// TwinCAT 3 PLC project TwinCAT_OpenFramework_HowTo
// Title: TwinCAT Open Framework HowTo
// Company: Oleksandr Tiutyk FOP
// Author: Oleksandr Tiutyk
// ProjectVersion: 1.0.13.0
// Description: Small samples how to use TwinCAT.OpenFramework
// ProgramVersion: 3.1.4026.28
// libraries:
//   [TwinCAT Open Framework Testing], * (Oleksandr Tiutyk FOP)
//   [TwinCAT Open Framework Core], * (Oleksandr Tiutyk FOP)
//   [TwinCAT Open Framework IO Models], * (Oleksandr Tiutyk FOP)
//   Tc2_Standard, * (Beckhoff Automation GmbH)
//   Tc2_System, * (Beckhoff Automation GmbH)
// project tree:
//   / CurrentNamespace.TcGVL, MAIN.TcPOU, PlcTask.TcTTO
//   Testing/ AdditionTestRunner.TcPOU, BasicTestRunner.TcPOU, TimerDelayTestRunner.TcPOU, AdditionTest.TcPOU, TimerDelayTest.TcPOU, SingleCycleTestExample.TcPOU, MultiCycleTestExample.TcPOU, TimingTestGroup.TcPOU, BasicTestGroup.TcPOU, GroupedTestExample.TcPOU
//   IO/ IOModelsExample.TcPOU
//   Version/ Global_Version.TcGVL
// (motion and I/O tree: see PLC project twincat_openframework_core)
// real-time tasks:
//   TASK PlcTask: cycle T#10ms, priority 20, ADS port 350
//   TASK TestTask: cycle T#10ms, priority 1, ADS port 351
//   TASK RunnerTestTask: cycle T#10ms, priority 2, ADS port 354
//   TASK HowToTask: cycle T#10ms, priority 22, ADS port 353
// variable links:

CONFIGURATION TwinCAT_OpenFramework_HowTo
    RESOURCE PLC ON TwinCAT3
        TASK PlcTask(INTERVAL := T#10ms, PRIORITY := 22);
        PROGRAM MAIN WITH PlcTask : MAIN;
    END_RESOURCE
END_CONFIGURATION

// ---- CurrentNamespace.TcGVL
(*
SPDX-FileCopyrightText: © 2026 Oleksandr Tiutyk <trofimich@gmail.com>
SPDX-License-Identifier: MIT
License: https://opensource.org/license/mit
*)

{attribute 'qualified_only'}
VAR_GLOBAL
	Name : STRING := 'TOF_Tests';
END_VAR

// ---- Version/Global_Version.TcGVL
{attribute 'TcGenerated'}
{attribute 'no-analysis'}
{attribute 'linkalways'}
// This function has been automatically generated from the project information.
VAR_GLOBAL CONSTANT
	{attribute 'const_non_replaced'}
	stLibVersion_TwinCAT_Open_Framework_HowTo : ST_LibVersion := (iMajor := 1, iMinor := 0, iBuild := 13, iRevision := 0, nFlags := 0, sVersion := '1.0.13.0');
END_VAR

// ---- MAIN.TcPOU
(*
SPDX-FileCopyrightText: © 2026 Oleksandr Tiutyk <trofimich@gmail.com>
SPDX-License-Identifier: MIT
License: https://opensource.org/license/mit
*)

(*!
<summary>Runs the standalone single-cycle testing example through its explicit execution method.</summary>
<description>Mapped by PlcTask. Do not also map SingleCycleTestExample to a task while this entry is used.</description>
*)

{attribute 'no_explicit_call' := 'do not call this function block directly'}
PROGRAM MAIN
VAR
	{attribute 'hide'}
	_ClassName : STRING := __POUNAME();
END_VAR

SingleCycleTestExample.Execute();

(*!
<summary>Borrows the concrete program name for its lifetime.</summary>
<description>Borrowed read-only storage; callers must not modify it.</description>
*)
{attribute 'monitoring' := 'call'}
PROPERTY ClassName : REFERENCE TO STRING
GET
ClassName REF= _ClassName;
END_GET
END_PROPERTY

(*!
<summary>Borrows the project namespace for the program lifetime.</summary>
<description>Borrowed read-only storage; callers must not modify it.</description>
*)
{attribute 'monitoring' := 'call'}
PROPERTY NamespaceName : REFERENCE TO STRING
GET
NamespaceName REF= CurrentNamespace.Name;
END_GET
END_PROPERTY

END_PROGRAM

// ---- Testing/SingleCycleTestExample.TcPOU
(*
SPDX-FileCopyrightText: © 2026 Oleksandr Tiutyk <trofimich@gmail.com>
SPDX-License-Identifier: MIT
License: https://opensource.org/license/mit
*)

(*!
<summary>Runs one single-cycle test directly, without a group.</summary>
<description>
Map this program to one cyclic PLC task or call its Execute method once per cycle from that task.
The concrete runner owns the tests; the program owns the reporter and performs task
cleanup at the end of every scan. Inspect _Runner.IsFinished, AllPassed and counts, then _Report.IsReady.
For independent task execution, assign SingleCycleTestExample and MultiCycleTestExample to different tasks.
They share no instances or mutable buffers. Do not assign the same program instance to multiple tasks.
</description>
*)

{attribute 'no_explicit_call' := 'do not call this function block directly'}
PROGRAM SingleCycleTestExample
VAR
	{attribute 'hide'}
	_ClassName : STRING := __POUNAME();

	_Runner : AdditionTestRunner;
	_Report : TOF_Testing.JUnitXmlReporter;
	_Configured : BOOL;
END_VAR

Execute();

//! <summary>Borrows the concrete program name for its lifetime; callers must not modify it.</summary>
{attribute 'monitoring' := 'call'}
PROPERTY ClassName : REFERENCE TO STRING
GET
ClassName REF= _ClassName;
END_GET
END_PROPERTY

(*!
<summary>Advances this example and performs standalone task-boundary memory cleanup.</summary>
<description>
Call once per cycle from the owning task, either through this method or by mapping this PROGRAM to that task.
Do not drive both entry paths or share the instance between tasks. Use as the standalone example in its task;
hosts with additional transient-exception consumers must provide a shared boundary instead.
</description>
*)
METHOD Execute
IF NOT _Configured THEN
	_Runner.Reporter := _Report;
	_Configured := TRUE;
END_IF

_Runner.Execute(cleanupTaskMemory := TRUE);
END_METHOD

(*!
<summary>Provides the library namespace used in diagnostics.</summary>
<description>
Borrowed read-only reference to the compiler-initialized library namespace; no ownership transfer.
</description>
*)
{attribute 'monitoring' := 'call'}
PROPERTY NamespaceName : REFERENCE TO STRING
GET
NamespaceName REF= CurrentNamespace.Name;
END_GET
END_PROPERTY

END_PROGRAM

// ---- Testing/AdditionTestRunner.TcPOU
(*
SPDX-License-Identifier: MIT
License: https://opensource.org/license/mit
*)

(*!
<summary>Runs one owned addition test without a group.</summary>
<description>
Owns persistent root instances and fixed child storage. Use from one task without reentry.
Children borrows the same array for the instance lifetime. Root parents remain zero.
</description>
*)

{attribute 'no_assign'}
{attribute 'no_explicit_call' := 'do not call this function block directly'}
FUNCTION_BLOCK AdditionTestRunner EXTENDS TOF_Testing.TestRunner<1>
VAR_STAT
	//! <summary>Class name shared by instances of this concrete runner.</summary>
	{attribute 'hide'}
	_ClassName : STRING := __POUNAME();
END_VAR
VAR
	{attribute 'hide'}
	{attribute 'init_namespace'}
	_NamespaceName : STRING;
END_VAR
VAR_OUTPUT
	//! <summary>Owned root element used by this runner.</summary>
	Root : AdditionTest(name := "Addition", parent := 0);
END_VAR
VAR
	_Children : ARRAY [0.._ChildCount - 1] OF TOF_Testing.ITestElement :=
	[
		Root
	];
END_VAR

(*!
<summary>Borrows the concrete class name; callers must not modify the returned storage.</summary>
*)
{attribute 'monitoring' := 'call'}
PROPERTY ClassName : REFERENCE TO STRING
GET
ClassName REF= _ClassName;
END_GET
END_PROPERTY

(*!
<summary>Borrows the concrete namespace name for the instance lifetime; callers must not modify it.</summary>
*)
{attribute 'monitoring' := 'call'}
PROPERTY NamespaceName : REFERENCE TO STRING
GET
NamespaceName REF= _NamespaceName;
END_GET
END_PROPERTY

(*!
<summary>Reports the complete concrete instance size.</summary>
*)
{attribute 'monitoring' := 'call'}
PROPERTY SelfSize : ULINT
GET
SelfSize := XSIZEOF(THIS^);
END_GET
END_PROPERTY

(*!
<summary>Borrows the unchanged persistent root array; application code must not modify it.</summary>
*)
{attribute 'monitoring' := 'call'}
PROPERTY Children : REFERENCE TO ARRAY [0.._ChildCount - 1] OF TOF_Testing.ITestElement
GET
Children REF= _Children;
END_GET
END_PROPERTY

END_FUNCTION_BLOCK

// ---- Testing/AdditionTest.TcPOU
(*
SPDX-FileCopyrightText: © 2026 Oleksandr Tiutyk <trofimich@gmail.com>
SPDX-License-Identifier: MIT
License: https://opensource.org/license/mit
*)

(*!
<summary>Shows a complete single-cycle test body without guards or contexts.</summary>
*)

{attribute 'no_explicit_call' := 'do not call this function block directly'}
FUNCTION_BLOCK AdditionTest EXTENDS TOF_Testing.SingleCycleTest
VAR_STAT
	{attribute 'hide'}
	_ClassName : STRING := __POUNAME();
END_VAR

//! <summary>Borrows the concrete class name for the lifetime of this instance; callers must not modify it.</summary>
{attribute 'monitoring' := 'call'}
PROPERTY ClassName : REFERENCE TO STRING
GET
ClassName REF= _ClassName;
END_GET
END_PROPERTY

(*!
<summary>Checks an arithmetic result and completes automatically on return.</summary>
*)
METHOD PROTECTED ExecuteTest
Assert.ThatDInt(actual := 2 + 3).ToBe(expected := 5);
END_METHOD

//! <summary>Borrows the compiler-initialized namespace; callers must not modify the returned reference.</summary>
{attribute 'monitoring' := 'call'}
PROPERTY NamespaceName : REFERENCE TO STRING
GET
NamespaceName REF= CurrentNamespace.Name;
END_GET
END_PROPERTY

//! <summary>Reports the complete concrete instance size, excluding separately allocated storage.</summary>
{attribute 'monitoring' := 'call'}
PROPERTY SelfSize : ULINT
GET
SelfSize := XSIZEOF(THIS^);
END_GET
END_PROPERTY

END_FUNCTION_BLOCK

// ---- Testing/BasicTestRunner.TcPOU
(*
SPDX-License-Identifier: MIT
License: https://opensource.org/license/mit
*)

(*!
<summary>Runs the owned basic test group and its nested timing group.</summary>
<description>
Owns persistent root instances and fixed child storage. Use from one task without reentry.
Children borrows the same array for the instance lifetime. Root parents remain zero.
</description>
*)

{attribute 'no_assign'}
{attribute 'no_explicit_call' := 'do not call this function block directly'}
FUNCTION_BLOCK BasicTestRunner EXTENDS TOF_Testing.TestRunner<1>
VAR_STAT
	//! <summary>Class name shared by instances of this concrete runner.</summary>
	{attribute 'hide'}
	_ClassName : STRING := __POUNAME();
END_VAR
VAR
	{attribute 'hide'}
	{attribute 'init_namespace'}
	_NamespaceName : STRING;
END_VAR
VAR_OUTPUT
	//! <summary>Owned root element used by this runner.</summary>
	Root : BasicTestGroup(name := "Basic", parent := 0);
END_VAR
VAR
	_Children : ARRAY [0.._ChildCount - 1] OF TOF_Testing.ITestElement :=
	[
		Root
	];
END_VAR

(*!
<summary>Borrows the concrete class name; callers must not modify the returned storage.</summary>
*)
{attribute 'monitoring' := 'call'}
PROPERTY ClassName : REFERENCE TO STRING
GET
ClassName REF= _ClassName;
END_GET
END_PROPERTY

(*!
<summary>Borrows the concrete namespace name for the instance lifetime; callers must not modify it.</summary>
*)
{attribute 'monitoring' := 'call'}
PROPERTY NamespaceName : REFERENCE TO STRING
GET
NamespaceName REF= _NamespaceName;
END_GET
END_PROPERTY

(*!
<summary>Reports the complete concrete instance size.</summary>
*)
{attribute 'monitoring' := 'call'}
PROPERTY SelfSize : ULINT
GET
SelfSize := XSIZEOF(THIS^);
END_GET
END_PROPERTY

(*!
<summary>Borrows the unchanged persistent root array; application code must not modify it.</summary>
*)
{attribute 'monitoring' := 'call'}
PROPERTY Children : REFERENCE TO ARRAY [0.._ChildCount - 1] OF TOF_Testing.ITestElement
GET
Children REF= _Children;
END_GET
END_PROPERTY

END_FUNCTION_BLOCK

// ---- Testing/BasicTestGroup.TcPOU
(*
SPDX-License-Identifier: MIT
License: https://opensource.org/license/mit
*)

(*!
<summary>Owns an arithmetic test and a nested timing group.</summary>
<description>
Owns persistent child storage and fixed parent associations. Use in one task without reentry.
Children is borrowed and must not be modified by application code. Constructor callbacks are not used.
</description>
*)

{attribute 'no_assign'}
{attribute 'no_explicit_call' := 'do not call this function block directly'}
FUNCTION_BLOCK BasicTestGroup EXTENDS TOF_Testing.TestGroup<2>
VAR_STAT
	{attribute 'hide'}
	_ClassName : STRING := __POUNAME();
END_VAR
VAR
	_Addition : AdditionTest(name := "Addition", parent := THIS^);
	_Timing : TimingTestGroup(name := "Timing", parent := THIS^);

	_Children : ARRAY [0.._ChildCount - 1] OF TOF_Testing.ITestElement :=
	[
		_Addition,
		_Timing
	];
END_VAR

//! <summary>Borrows the fixed array of this concrete group; do not modify it.</summary>
{attribute 'monitoring' := 'call'}
PROPERTY Children : REFERENCE TO ARRAY [0.._ChildCount - 1] OF TOF_Testing.ITestElement
GET
Children REF= _Children;
END_GET
END_PROPERTY

//! <summary>Borrows the concrete class name for the lifetime of this instance; callers must not modify it.</summary>
{attribute 'monitoring' := 'call'}
PROPERTY ClassName : REFERENCE TO STRING
GET
ClassName REF= _ClassName;
END_GET
END_PROPERTY

//! <summary>Borrows the compiler-initialized namespace; callers must not modify the returned reference.</summary>
{attribute 'monitoring' := 'call'}
PROPERTY NamespaceName : REFERENCE TO STRING
GET
NamespaceName REF= CurrentNamespace.Name;
END_GET
END_PROPERTY

//! <summary>Reports the complete concrete instance size, excluding separately allocated storage.</summary>
{attribute 'monitoring' := 'call'}
PROPERTY SelfSize : ULINT
GET
SelfSize := XSIZEOF(THIS^);
END_GET
END_PROPERTY

END_FUNCTION_BLOCK

// ---- Testing/TimingTestGroup.TcPOU
(*
SPDX-License-Identifier: MIT
License: https://opensource.org/license/mit
*)

(*!
<summary>Owns a timer-delay test as a static group.</summary>
<description>
Owns persistent child storage and fixed parent associations. Use in one task without reentry.
Children is borrowed and must not be modified by application code. Constructor callbacks are not used.
</description>
*)

{attribute 'no_assign'}
{attribute 'no_explicit_call' := 'do not call this function block directly'}
FUNCTION_BLOCK TimingTestGroup EXTENDS TOF_Testing.TestGroup<1>
VAR_STAT
	//! <summary>Class name shared by all instances of this function block.</summary>
	{attribute 'hide'}
	_ClassName : STRING := __POUNAME();
END_VAR
VAR
	_Timer : TimerDelayTest(name := "Timer delay", parent := THIS^);

	_Children : ARRAY [0.._ChildCount - 1] OF TOF_Testing.ITestElement :=
	[
		_Timer
	];
END_VAR

//! <summary>Borrows the fixed array of this concrete group; do not modify it.</summary>
{attribute 'monitoring' := 'call'}
PROPERTY Children : REFERENCE TO ARRAY [0.._ChildCount - 1] OF TOF_Testing.ITestElement
GET
Children REF= _Children;
END_GET
END_PROPERTY

//! <summary>Borrows the concrete class name for the lifetime of this instance; callers must not modify it.</summary>
{attribute 'monitoring' := 'call'}
PROPERTY ClassName : REFERENCE TO STRING
GET
ClassName REF= _ClassName;
END_GET
END_PROPERTY

//! <summary>Borrows the compiler-initialized namespace; callers must not modify the returned reference.</summary>
{attribute 'monitoring' := 'call'}
PROPERTY NamespaceName : REFERENCE TO STRING
GET
NamespaceName REF= CurrentNamespace.Name;
END_GET
END_PROPERTY

//! <summary>Reports the complete concrete instance size, excluding separately allocated storage.</summary>
{attribute 'monitoring' := 'call'}
PROPERTY SelfSize : ULINT
GET
SelfSize := XSIZEOF(THIS^);
END_GET
END_PROPERTY

END_FUNCTION_BLOCK

// ---- Testing/TimerDelayTest.TcPOU
(*
SPDX-FileCopyrightText: © 2026 Oleksandr Tiutyk <trofimich@gmail.com>
SPDX-License-Identifier: MIT
License: https://opensource.org/license/mit
*)

(*!
<summary>Shows persistent state and explicit completion in a multi-cycle test.</summary>
<description>
The inherited one-second deadline bounds waiting for a twenty-millisecond timer.
</description>
*)

{attribute 'no_explicit_call' := 'do not call this function block directly'}
FUNCTION_BLOCK TimerDelayTest EXTENDS TOF_Testing.MultiCycleTest
VAR
	_Timer : Tc2_Standard.TON;
END_VAR
VAR_STAT
	//! <summary>Class name shared by all instances of this function block.</summary>
	{attribute 'hide'}
	_ClassName : STRING := __POUNAME();
END_VAR
VAR
	{attribute 'hide'}
	{attribute 'init_namespace'}
	_NamespaceName : STRING;
END_VAR

(*!
<summary>Resets the timer after completion or failure.</summary>
*)
METHOD PROTECTED AfterTest
_Timer(IN := FALSE, PT := T#20MS);
END_METHOD

(*!
<summary>Resets the timer before each run.</summary>
*)
METHOD PROTECTED BeforeTest
_Timer(IN := FALSE, PT := T#20MS);
END_METHOD

//! <summary>Borrows the concrete class name for the lifetime of this instance; callers must not modify it.</summary>
{attribute 'monitoring' := 'call'}
PROPERTY ClassName : REFERENCE TO STRING
GET
ClassName REF= _ClassName;
END_GET
END_PROPERTY

(*!
<summary>Advances the timer once and returns DONE after its delay.</summary>
*)
METHOD PROTECTED ExecuteTest : TOF_Testing.TEST_CYCLE_RESULT
_Timer(IN := TRUE, PT := T#20MS);

IF _Timer.Q THEN
	Assert.ThatTime(actual := _Timer.ET).IsGreaterThanOrEquals(expected := T#20MS);
	ExecuteTest := TOF_Testing.TEST_CYCLE_RESULT.DONE;
ELSE
	ExecuteTest := TOF_Testing.TEST_CYCLE_RESULT.BUSY;
END_IF
END_METHOD

//! <summary>Borrows the compiler-initialized namespace; callers must not modify the returned reference.</summary>
{attribute 'monitoring' := 'call'}
PROPERTY NamespaceName : REFERENCE TO STRING
GET
NamespaceName REF= CurrentNamespace.Name;
END_GET
END_PROPERTY

//! <summary>Reports the complete concrete instance size, excluding separately allocated storage.</summary>
{attribute 'monitoring' := 'call'}
PROPERTY SelfSize : ULINT
GET
SelfSize := XSIZEOF(THIS^);
END_GET
END_PROPERTY

END_FUNCTION_BLOCK

// ---- Testing/TimerDelayTestRunner.TcPOU
(*
SPDX-License-Identifier: MIT
License: https://opensource.org/license/mit
*)

(*!
<summary>Runs one owned multi-cycle timer test.</summary>
<description>
Owns persistent root instances and fixed child storage. Use from one task without reentry.
Children borrows the same array for the instance lifetime. Root parents remain zero.
</description>
*)

{attribute 'no_assign'}
{attribute 'no_explicit_call' := 'do not call this function block directly'}
FUNCTION_BLOCK TimerDelayTestRunner EXTENDS TOF_Testing.TestRunner<1>
VAR_STAT
	//! <summary>Class name shared by instances of this concrete runner.</summary>
	{attribute 'hide'}
	_ClassName : STRING := __POUNAME();
END_VAR
VAR
	{attribute 'hide'}
	{attribute 'init_namespace'}
	_NamespaceName : STRING;
END_VAR
VAR_OUTPUT
	//! <summary>Owned root element used by this runner.</summary>
	Root : TimerDelayTest(name := "Timer delay", parent := 0);
END_VAR
VAR
	_Children : ARRAY [0.._ChildCount - 1] OF TOF_Testing.ITestElement :=
	[
		Root
	];
END_VAR

(*!
<summary>Borrows the concrete class name; callers must not modify the returned storage.</summary>
*)
{attribute 'monitoring' := 'call'}
PROPERTY ClassName : REFERENCE TO STRING
GET
ClassName REF= _ClassName;
END_GET
END_PROPERTY

(*!
<summary>Borrows the concrete namespace name for the instance lifetime; callers must not modify it.</summary>
*)
{attribute 'monitoring' := 'call'}
PROPERTY NamespaceName : REFERENCE TO STRING
GET
NamespaceName REF= _NamespaceName;
END_GET
END_PROPERTY

(*!
<summary>Reports the complete concrete instance size.</summary>
*)
{attribute 'monitoring' := 'call'}
PROPERTY SelfSize : ULINT
GET
SelfSize := XSIZEOF(THIS^);
END_GET
END_PROPERTY

(*!
<summary>Borrows the unchanged persistent root array; application code must not modify it.</summary>
*)
{attribute 'monitoring' := 'call'}
PROPERTY Children : REFERENCE TO ARRAY [0.._ChildCount - 1] OF TOF_Testing.ITestElement
GET
Children REF= _Children;
END_GET
END_PROPERTY

END_FUNCTION_BLOCK

// ---- Testing/MultiCycleTestExample.TcPOU
(*
SPDX-FileCopyrightText: © 2026 Oleksandr Tiutyk <trofimich@gmail.com>
SPDX-License-Identifier: MIT
License: https://opensource.org/license/mit
*)

(*!
<summary>Runs one multi-cycle test until completion or the inherited deadline.</summary>
<description>
Map this program to one cyclic PLC task or call its Execute method once per cycle from that task.
The concrete runner owns the tests; the program owns the reporter and performs task
cleanup at the end of every scan. Inspect _Runner.IsFinished, AllPassed and counts, then _Report.IsReady.
For independent task execution, assign SingleCycleTestExample and MultiCycleTestExample to different tasks.
They share no instances or mutable buffers. Do not assign the same program instance to multiple tasks.
</description>
*)

{attribute 'no_explicit_call' := 'do not call this function block directly'}
PROGRAM MultiCycleTestExample
VAR
	{attribute 'hide'}
	_ClassName : STRING := __POUNAME();

	_Runner : TimerDelayTestRunner;
	_Report : TOF_Testing.JUnitXmlReporter;
	_Configured : BOOL;
END_VAR

Execute();

//! <summary>Borrows the concrete program name for its lifetime; callers must not modify it.</summary>
{attribute 'monitoring' := 'call'}
PROPERTY ClassName : REFERENCE TO STRING
GET
ClassName REF= _ClassName;
END_GET
END_PROPERTY

(*!
<summary>Advances this example and performs standalone task-boundary memory cleanup.</summary>
<description>
Call once per cycle from the owning task, either through this method or by mapping this PROGRAM to that task.
Do not drive both entry paths or share the instance between tasks. Use as the standalone example in its task;
hosts with additional transient-exception consumers must provide a shared boundary instead.
</description>
*)
METHOD Execute
IF NOT _Configured THEN
	_Runner.Reporter := _Report;
	_Configured := TRUE;
END_IF

_Runner.Execute(cleanupTaskMemory := TRUE);
END_METHOD

(*!
<summary>Provides the library namespace used in diagnostics.</summary>
<description>
Borrowed read-only reference to the compiler-initialized library namespace; no ownership transfer.
</description>
*)
{attribute 'monitoring' := 'call'}
PROPERTY NamespaceName : REFERENCE TO STRING
GET
NamespaceName REF= CurrentNamespace.Name;
END_GET
END_PROPERTY

END_PROGRAM

// ---- Testing/GroupedTestExample.TcPOU
(*
SPDX-FileCopyrightText: © 2026 Oleksandr Tiutyk <trofimich@gmail.com>
SPDX-License-Identifier: MIT
License: https://opensource.org/license/mit
*)

(*!
<summary>Runs a single-cycle and a multi-cycle test through nested sequential groups.</summary>
<description>
Map this program to one cyclic PLC task or call its Execute method once per cycle from that task.
The concrete runner owns the tests; the program owns the reporter and performs task
cleanup at the end of every scan. Inspect _Runner.IsFinished, AllPassed and counts, then _Report.IsReady.
For independent task execution, assign SingleCycleTestExample and MultiCycleTestExample to different tasks.
They share no instances or mutable buffers. Do not assign the same program instance to multiple tasks.
</description>
*)

{attribute 'no_explicit_call' := 'do not call this function block directly'}
PROGRAM GroupedTestExample
VAR
	{attribute 'hide'}
	_ClassName : STRING := __POUNAME();

	_Runner : BasicTestRunner;
	_Report : TOF_Testing.JUnitXmlReporter;
	_Configured : BOOL;
END_VAR

Execute();

//! <summary>Borrows the concrete program name for its lifetime; callers must not modify it.</summary>
{attribute 'monitoring' := 'call'}
PROPERTY ClassName : REFERENCE TO STRING
GET
ClassName REF= _ClassName;
END_GET
END_PROPERTY

(*!
<summary>Advances this example and performs standalone task-boundary memory cleanup.</summary>
<description>
Call once per cycle from the owning task, either through this method or by mapping this PROGRAM to that task.
Do not drive both entry paths or share the instance between tasks. Use as the standalone example in its task;
hosts with additional transient-exception consumers must provide a shared boundary instead.
</description>
*)
METHOD Execute
IF NOT _Configured THEN
	_Runner.Reporter := _Report;
	_Configured := TRUE;
END_IF

_Runner.Execute(cleanupTaskMemory := TRUE);
END_METHOD

(*!
<summary>Provides the library namespace used in diagnostics.</summary>
<description>
Borrowed read-only reference to the compiler-initialized library namespace; no ownership transfer.
</description>
*)
{attribute 'monitoring' := 'call'}
PROPERTY NamespaceName : REFERENCE TO STRING
GET
NamespaceName REF= CurrentNamespace.Name;
END_GET
END_PROPERTY

END_PROGRAM

// ---- IO/IOModelsExample.TcPOU
(*
SPDX-FileCopyrightText: © 2026 Oleksandr Tiutyk <trofimich@gmail.com>
SPDX-License-Identifier: MIT
License: https://opensource.org/license/mit
*)

(*!
<summary>Demonstrates explicit EL3001 mapping, input validity and update observation without a test framework.</summary>
<description>
Select the EL3001 standard status-plus-INT16 PDO. Link _Terminal.Ch1.Status and Value, WcState, InputToggle,
State and AdsAddr to the corresponding slave entries in XAE, then set BindingsConfigured to TRUE.
The flag records caller confirmation; software cannot detect unlinked zero-valued inputs.
Map this program to one task or call Execute once per cycle from that task. Use only one execution path.
Voltage is zero while InputValid is FALSE; use InputValid before consuming Voltage. InputUpdated observes
a toggle transition, not the level of InputToggle. State and AdsAddr are acyclic and do not validate measurements.
The program owns no dynamic resources. Execute checks the fatal allocation latch outside recoverable handlers;
a hosting task remains responsible for cleanup after all of its transient-exception consumers.
Do not copy the program or share its mutable state across tasks without external synchronization.
</description>
*)

{attribute 'no_explicit_call' := 'do not call this function block directly'}
PROGRAM IOModelsExample
VAR CONSTANT
	//! <summary>Positive full-scale signed raw code used for the EL3001 voltage scaling.</summary>
	_FullScaleRawValue : LREAL := 32767.0;
	//! <summary>Positive electrical full scale of the selected EL3001 range, in volts.</summary>
	_FullScaleVoltage : LREAL := 10.0;
END_VAR
VAR
	_ClassName : STRING := __POUNAME();
	_Terminal : TOF_IOModels.EL3001_EX;
	_BindingsConfigured : BOOL;
	_InputValid : BOOL;
	_InputUpdated : BOOL;
	_PreviousToggle : BOOL;
	_Voltage : LREAL;
END_VAR

Execute();

(*!
<summary>Samples the configured input and exposes guarded voltage and update observations.</summary>
<description>
Call once per scan from the owning task. Reading mapped fields is not an atomic cross-task snapshot.
Fatal allocation failure propagates at this task boundary; no handler here can convert it into normal operation.
</description>
*)
METHOD Execute
TOF_Core.DynamicMemoryManager.RaiseIfAllocationFailed();

_InputValid := _BindingsConfigured
	AND_THEN NOT _Terminal.WcState
	AND_THEN NOT _Terminal.Ch1.Status.6
	AND_THEN NOT _Terminal.Ch1.Status.14;
_InputUpdated := _InputValid AND_THEN (_Terminal.InputToggle <> _PreviousToggle);
_PreviousToggle := _Terminal.InputToggle;

IF _InputValid THEN
	_Voltage := TO_LREAL(_Terminal.Ch1.Value) * _FullScaleVoltage / _FullScaleRawValue;
ELSE
	_Voltage := 0.0;
END_IF
END_METHOD

(*!
<summary>Records caller confirmation that all required XAE links and the selected PDO are configured.</summary>
<description>Set TRUE only after mapping inspection. FALSE inhibits measurement use on the next Execute.</description>
*)
PROPERTY BindingsConfigured : BOOL
GET
BindingsConfigured := _BindingsConfigured;
END_GET
SET
_BindingsConfigured := BindingsConfigured;
END_SET
END_PROPERTY

//! <summary>Reports the bus/channel validity evaluated during the latest Execute.</summary>
PROPERTY InputValid : BOOL
GET
InputValid := _InputValid;
END_GET
END_PROPERTY

//! <summary>Reports a valid input-toggle transition observed during the latest Execute.</summary>
PROPERTY InputUpdated : BOOL
GET
InputUpdated := _InputUpdated;
END_GET
END_PROPERTY

(*!
<summary>Returns the latest guarded EL3001 voltage in volts.</summary>
<description>Zero while InputValid is FALSE; inspect InputValid because a valid voltage can also be zero.</description>
*)
PROPERTY Voltage : LREAL
GET
Voltage := _Voltage;
END_GET
END_PROPERTY

//! <summary>Borrows the program-owned concrete name; callers must not modify it.</summary>
PROPERTY ClassName : REFERENCE TO STRING
GET
ClassName REF= _ClassName;
END_GET
END_PROPERTY

//! <summary>Borrows project namespace storage for the program lifetime; callers must not modify it.</summary>
PROPERTY NamespaceName : REFERENCE TO STRING
GET
NamespaceName REF= CurrentNamespace.Name;
END_GET
END_PROPERTY

END_PROGRAM
